{attribute 'namespace' := 'MyLib.Modbus'}
TYPE eMbCycleState :
(
    eMbState_Init,
    eMbState_Read,
    eMbState_Write,
    eMbState_Error
);
END_TYPE

(* stored: Version 1.1.0.1, ProductVersion 3.1.4024.13
   DUT eMbCycleState: Id {ca6d863a-a1cb-4128-a8c2-f50894e8cd56} *)
